(* IEC 61131-3 sources: rusty/tests/lit/single/type_promotion/for_loop, 9 files *)

(* ---- step_evaluated_once_per_iteration.st ---- *)
// RUN: %COMPILE %s && %RUN | %CHECK %s
// The step is evaluated once per iteration, so the counter value that the loop tests is the value that the body sees.
VAR_GLOBAL
    calls : DINT;
    step : DINT;
END_VAR

FUNCTION next_step : DINT
    calls := calls + 1;
    next_step := calls;
END_FUNCTION

FUNCTION end_changes_step : DINT
    step := step + 1;
    end_changes_step := 2;
END_FUNCTION

FUNCTION main : DINT
    VAR
        i : DINT;
    END_VAR

    // The direction test reads 1, then the passes read 2 and 3
    calls := 0;
    FOR i := 0 TO 2 BY next_step() DO
        printf('BY next_step(): i = %d$N', i);
    END_FOR
    printf('BY next_step(): after = %d, calls = %d$N', i, calls);
    // CHECK:      BY next_step(): i = 0
    // CHECK-NEXT: BY next_step(): i = 2
    // CHECK-NEXT: BY next_step(): after = 5, calls = 3

    // The end value changes the step after the step is read
    step := 1;
    FOR i := 0 TO end_changes_step() BY step DO
        printf('TO end_changes_step(): i = %d$N', i);
    END_FOR
    printf('TO end_changes_step(): after = %d$N', i);
    // CHECK-NEXT: TO end_changes_step(): i = 0
    // CHECK-NEXT: TO end_changes_step(): i = 2
    // CHECK-NEXT: TO end_changes_step(): after = 5
END_FUNCTION

(* ---- counter_types.st ---- *)
// RUN: %COMPILE %s && %RUN | %CHECK %s
// The next counter value is a LINT for an integer, bit-string or BOOL counter of up to 32 bits, and has the counter's
// own type otherwise, so every counter type ends at its end value.
FUNCTION other : DINT
    VAR
        __next_0 : LREAL;
        r : REAL := 1.5;
    END_VAR
    // A user variable with the name of a loop temporary does not change the loop
    __next_0 := r;
    other := 0;
END_FUNCTION

FUNCTION main : DINT
    VAR
        d : DINT;
        ud : UDINT;
        b : BOOL;
        t : TIME;
        r : REAL;
        ul : ULINT;
        n : DINT;
        after : LINT;
    END_VAR

    n := 0;
    FOR d := 16777216 TO 16777220 DO
        n := n + 1;
        IF n > 100 THEN EXIT; END_IF
    END_FOR
    printf('DINT 16777216 TO 16777220 = %d$N', n);                                   // CHECK: DINT 16777216 TO 16777220 = 5

    n := 0;
    FOR ud := 2400000000 TO 2000000000 BY -100000000 DO
        n := n + 1;
        IF n > 100 THEN EXIT; END_IF
    END_FOR
    after := ud;
    printf('UDINT 2400000000 TO 2000000000 BY -100000000 = %d, after = %lld$N', n, after);
    // CHECK-NEXT: UDINT 2400000000 TO 2000000000 BY -100000000 = 5, after = 1900000000

    n := 0;
    FOR b := FALSE TO TRUE DO
        n := n + 1;
        IF n > 100 THEN EXIT; END_IF
    END_FOR
    printf('BOOL FALSE TO TRUE = %d$N', n);                                          // CHECK-NEXT: BOOL FALSE TO TRUE = 2

    n := 0;
    FOR t := T#1s TO T#3s BY T#1s DO
        n := n + 1;
        IF n > 100 THEN EXIT; END_IF
    END_FOR
    printf('TIME T#1s TO T#3s BY T#1s = %d$N', n);                                   // CHECK-NEXT: TIME T#1s TO T#3s BY T#1s = 3

    n := 0;
    FOR r := 0.0 TO 1.0 BY 0.25 DO
        n := n + 1;
        IF n > 100 THEN EXIT; END_IF
    END_FOR
    printf('REAL 0.0 TO 1.0 BY 0.25 = %d, after = %.2f$N', n, r);                    // CHECK-NEXT: REAL 0.0 TO 1.0 BY 0.25 = 5, after = 1.25

    n := 0;
    FOR ul := 9223372036854775806 TO 9223372036854775810 DO
        n := n + 1;
        IF n > 100 THEN EXIT; END_IF
    END_FOR
    printf('ULINT across 2^63 = %d$N', n);                                           // CHECK-NEXT: ULINT across 2^63 = 5
END_FUNCTION

(* ---- counter_with_64_bit_end.st ---- *)
// RUN: %COMPILE %s && %RUN | %CHECK %s
// A counter narrower than 64 bits with a LINT or ULINT end value runs the expected number of passes.
FUNCTION main : DINT
    VAR
        us : USINT;
        ud : UDINT;
        d : DINT;
        end_l : LINT := 5;
        end_ul : ULINT := 5;
        step : SINT := 2;
        n : DINT;
    END_VAR

    n := 0;
    FOR us := 1 TO end_l DO
        n := n + 1;
        IF n > 1000 THEN EXIT; END_IF
    END_FOR
    printf('USINT 1 TO LINT 5 = %d$N', n);                      // CHECK: USINT 1 TO LINT 5 = 5

    n := 0;
    FOR ud := 1 TO end_ul DO
        n := n + 1;
        IF n > 1000 THEN EXIT; END_IF
    END_FOR
    printf('UDINT 1 TO ULINT 5 = %d$N', n);                     // CHECK-NEXT: UDINT 1 TO ULINT 5 = 5

    n := 0;
    FOR d := 1 TO end_l BY step DO
        n := n + 1;
        IF n > 1000 THEN EXIT; END_IF
    END_FOR
    printf('DINT 1 TO LINT 5 BY SINT 2 = %d$N', n);             // CHECK-NEXT: DINT 1 TO LINT 5 BY SINT 2 = 3
END_FUNCTION

(* ---- counter_within_type_range.st ---- *)
// RUN: %COMPILE %s && %RUN | %CHECK %s
// FOR loops whose counter stays inside the range of its type.
FUNCTION main : DINT
    VAR
        us : USINT;
        ud : UDINT;
        s : SINT;
        n : DINT;
    END_VAR

    n := 0;
    FOR us := 1 TO 10 BY 3 DO
        n := n + 1;
    END_FOR
    printf('USINT 1 TO 10 BY 3 = %d$N', n);                 // CHECK: USINT 1 TO 10 BY 3 = 4

    n := 0;
    FOR us := 10 TO 1 BY -1 DO
        n := n + 1;
    END_FOR
    printf('USINT 10 TO 1 BY -1 = %d$N', n);                // CHECK-NEXT: USINT 10 TO 1 BY -1 = 10

    n := 0;
    FOR us := 200 TO 220 BY 10 DO
        n := n + 1;
    END_FOR
    printf('USINT 200 TO 220 BY 10 = %d$N', n);             // CHECK-NEXT: USINT 200 TO 220 BY 10 = 3

    n := 0;
    FOR ud := 10 TO 1 BY -3 DO
        n := n + 1;
    END_FOR
    printf('UDINT 10 TO 1 BY -3 = %d$N', n);                // CHECK-NEXT: UDINT 10 TO 1 BY -3 = 4

    n := 0;
    FOR s := 10 TO -10 BY -5 DO
        n := n + 1;
    END_FOR
    printf('SINT 10 TO -10 BY -5 = %d$N', n);               // CHECK-NEXT: SINT 10 TO -10 BY -5 = 5
END_FUNCTION

(* ---- counter_wraps_past_64_bit_limit.st ---- *)
// RUN: %COMPILE %s && %RUN | %CHECK %s
// XFAIL: *
// For a 64-bit counter, the next value has the counter's own type, so a next value past the type's limit wraps before the end test and the loop goes on.
FUNCTION main : DINT
    VAR
        ul : ULINT;
        l : LINT;
        n : DINT;
    END_VAR

    n := 0;
    FOR ul := 10 TO 0 BY -1 DO
        n := n + 1;
        IF n > 1000 THEN EXIT; END_IF
    END_FOR
    printf('ULINT 10 TO 0 BY -1 = %d$N', n);                                    // CHECK: ULINT 10 TO 0 BY -1 = 11

    n := 0;
    FOR l := 9223372036854775800 TO 9223372036854775807 BY 5 DO
        n := n + 1;
        IF n > 1000 THEN EXIT; END_IF
    END_FOR
    printf('LINT 9223372036854775800 TO 9223372036854775807 BY 5 = %d$N', n);  // CHECK-NEXT: LINT 9223372036854775800 TO 9223372036854775807 BY 5 = 2
END_FUNCTION

(* ---- counter_wraps_past_type_limit.st ---- *)
// RUN: %COMPILE %s && %RUN | %CHECK %s
// A next value past the limit of a counter of up to 32 bits ends the loop. The counter keeps the wrapped value.
FUNCTION main : DINT
    VAR
        us : USINT;
        s : SINT;
        bt : BYTE;
        ud : UDINT;
        d : DINT;
        step : SINT;
        n : DINT;
        after : LINT;
    END_VAR

    // Below the minimum
    n := 0;
    FOR us := 10 TO 1 BY -3 DO
        n := n + 1;
        IF n > 1000 THEN EXIT; END_IF
    END_FOR
    after := us;
    printf('USINT 10 TO 1 BY -3 = %d, after = %lld$N', n, after);
    // CHECK: USINT 10 TO 1 BY -3 = 4, after = 254

    n := 0;
    FOR ud := 5 TO 0 BY -2 DO
        n := n + 1;
        IF n > 1000 THEN EXIT; END_IF
    END_FOR
    after := ud;
    printf('UDINT 5 TO 0 BY -2 = %d, after = %lld$N', n, after);
    // CHECK-NEXT: UDINT 5 TO 0 BY -2 = 3, after = 4294967295

    // Past the maximum
    n := 0;
    FOR s := 120 TO 127 BY 5 DO
        n := n + 1;
        IF n > 1000 THEN EXIT; END_IF
    END_FOR
    after := s;
    printf('SINT 120 TO 127 BY 5 = %d, after = %lld$N', n, after);
    // CHECK-NEXT: SINT 120 TO 127 BY 5 = 2, after = -126

    n := 0;
    FOR d := 2147483640 TO 2147483647 BY 5 DO
        n := n + 1;
        IF n > 1000 THEN EXIT; END_IF
    END_FOR
    after := d;
    printf('DINT 2147483640 TO 2147483647 BY 5 = %d, after = %lld$N', n, after);
    // CHECK-NEXT: DINT 2147483640 TO 2147483647 BY 5 = 2, after = -2147483646

    n := 0;
    FOR bt := 250 TO 255 BY BYTE#3 DO
        n := n + 1;
        IF n > 1000 THEN EXIT; END_IF
    END_FOR
    after := bt;
    printf('BYTE 250 TO 255 BY BYTE#3 = %d, after = %lld$N', n, after);
    // CHECK-NEXT: BYTE 250 TO 255 BY BYTE#3 = 2, after = 0

    // A step larger than the counter's range
    n := 0;
    FOR us := 10 TO 200 BY 300 DO
        n := n + 1;
        IF n > 1000 THEN EXIT; END_IF
    END_FOR
    after := us;
    printf('USINT 10 TO 200 BY 300 = %d, after = %lld$N', n, after);
    // CHECK-NEXT: USINT 10 TO 200 BY 300 = 1, after = 54

    // CONTINUE does not skip the end test
    n := 0;
    FOR us := 250 TO 255 BY 3 DO
        n := n + 1;
        IF n > 1000 THEN EXIT; END_IF
        CONTINUE;
    END_FOR
    after := us;
    printf('USINT 250 TO 255 BY 3 with CONTINUE = %d, after = %lld$N', n, after);
    // CHECK-NEXT: USINT 250 TO 255 BY 3 with CONTINUE = 2, after = 0

    // A step changed in the body moves the counter past the limit
    n := 0;
    step := 1;
    FOR us := 250 TO 255 BY step DO
        n := n + 1;
        step := 4;
        IF n > 1000 THEN EXIT; END_IF
    END_FOR
    after := us;
    printf('USINT 250 TO 255 BY step = %d, after = %lld$N', n, after);
    // CHECK-NEXT: USINT 250 TO 255 BY step = 2, after = 2
END_FUNCTION

(* ---- date_counter_with_time_step.st ---- *)
// RUN: not %COMPILE --error-format clang %s 2>&1 | %CHECK %s
// A DATE counter computes its next value as a DATE, so a TIME step is an error, as in `d + T#1d`.
FUNCTION main : DINT
    VAR
        d : DATE;
        n : DINT;
    END_VAR

    FOR d := D#2020-01-01 TO D#2020-01-05 BY T#1d DO
        n := n + 1;
    END_FOR
END_FUNCTION

// CHECK: error[E156]: Operator `+` is not defined for `DATE` and `TIME`

(* ---- parenthesized_step.st ---- *)
// RUN: %COMPILE %s && %RUN | %CHECK %s
// A step in parentheses gives the same number of passes as without parentheses.
FUNCTION main : DINT
    VAR
        ul : ULINT;
        lw : LWORD;
        step : SINT := 2;
        n : DINT;
    END_VAR

    n := 0;
    FOR ul := 1 TO 7 BY (step) DO
        n := n + 1;
        IF n > 1000 THEN EXIT; END_IF
    END_FOR
    printf('ULINT 1 TO 7 BY (step) = %d$N', n);         // CHECK: ULINT 1 TO 7 BY (step) = 4

    n := 0;
    FOR lw := 1 TO 7 BY ((step)) DO
        n := n + 1;
        IF n > 1000 THEN EXIT; END_IF
    END_FOR
    printf('LWORD 1 TO 7 BY ((step)) = %d$N', n);       // CHECK-NEXT: LWORD 1 TO 7 BY ((step)) = 4
END_FUNCTION

(* ---- warnings_of_the_end_test.st ---- *)
// RUN: %COMPILE %s --error-format clang 2>&1 | %CHECK %s
// A FOR loop reports the operand conversion warnings of its end test `<next value> > <end>` (or `<`). The next
// value is a LINT for a counter of up to 32 bits and has the counter's type otherwise. The other generated
// statements report none.

FUNCTION main : DINT
    VAR
        c_int : INT;
        c_udint : UDINT;
        c_ulint : ULINT;
        c_lword : LWORD;
        step : DINT;
        end_d : DINT;
        end_u : UDINT;
        end_l : LINT;
        end_ul : ULINT;
        end_r : REAL;
    END_VAR

    // CHECK-NOT: {{.*}}warning{{.*}}
    FOR c_int := 10 TO 1 BY -3 DO END_FOR
    FOR c_int := 1 TO end_u BY step DO END_FOR
    FOR c_udint := 1 TO end_d DO END_FOR
    // CHECK: {{.*}}.st:[[@LINE+1]]:25:{{.*}}: warning[E161]: Operand of type 'ULINT' is converted to 'LINT', which may change its sign.
    FOR c_udint := 1 TO end_ul DO END_FOR
    // CHECK-NEXT: {{.*}}.st:[[@LINE+1]]:25:{{.*}}: warning[E161]: Operand of type 'DINT' is converted to 'ULINT', which may change its sign.
    FOR c_ulint := 1 TO end_d DO END_FOR
    // CHECK-NEXT: {{.*}}.st:[[@LINE+1]]:9:{{.*}}: warning[E161]: Operand of type 'ULINT' is converted to 'LINT', which may change its sign.
    FOR c_ulint := 1 TO end_l DO END_FOR
    // CHECK-NEXT: {{.*}}.st:[[@LINE+1]]:9:{{.*}}: warning[E161]: Operand of type 'LWORD' is converted to 'LINT', which may change its sign.
    FOR c_lword := 1 TO end_l BY step DO END_FOR
    // CHECK-NEXT: {{.*}}.st:[[@LINE+1]]:9:{{.*}}: warning[E162]: Implicit conversion from 'LINT' to 'LREAL' may lose precision.
    FOR c_int := 1 TO end_r DO END_FOR
END_FUNCTION

// CHECK-NOT: {{.*}}warning{{.*}}
